// TIA Portal V20 export
// export: Created 2026-10-11T05:31:09.1029328Z, ExportSetting WithDefaults, DisplayName Totally Integrated Automation Portal, DisplayVersion V20, DisplayName TIA Portal Openness, DisplayVersion V20, DisplayName TIA Portal Teamcenter Gateway, DisplayVersion V20, DisplayName TIA Portal Version Control Interface, DisplayVersion V20, DisplayName SINAMICS Startdrive Advanced, DisplayVersion V20 SP1 Update 2, DisplayName SINAMICS Startdrive G110M, G120, G120C, G120D, G120P, G115D, DisplayVersion V20 SP1 Update 2, DisplayName SINAMICS Startdrive G130, G150, S120, S150, SINAMICS MV, G220, S200, S210, DisplayVersion V20 SP1 Update 2, DisplayName STEP 7 Professional, DisplayVersion V20, DisplayName STEP 7 Safety, DisplayVersion V20, DisplayName WinCC Basic/Comfort/Advanced, DisplayVersion V20, DisplayName WinCC Professional, DisplayVersion V20, DisplayName WinCC Unified, DisplayVersion V20
FUNCTION "FRK_UnitMode" : Void   // FC47, SCL
{ S7_Optimized_Access := 'TRUE' }
VERSION : 0.1
// stored: AutoNumber true, IsIECCheckEnabled false, SetENOAutomatically false, UDAEnableTagReadback false
   VAR_IN_OUT
      Core : "FRK_Core";
      Unit : "FRK_Unit";
   END_VAR
BEGIN

   IF #Unit.ModePending THEN
       IF #Core.Exec = 1 THEN
           #Core.EvModeExit := TRUE;
           #Core.HookResult := 0;
       ELSIF #Core.Exec = 0 AND NOT #Unit.Clearing THEN
           #Unit.Mode := #Unit.RequestedMode;
           #Unit.ModePending := FALSE;
           #Unit.ExitFirst := FALSE;
           #Core.EvModeChanged := TRUE;
       ELSE
           #Unit.RunReq := FALSE;
       END_IF;
   END_IF;
END_FUNCTION
